(* IEC 61131-3 sources: esbmc-plc-benchmark-suite/ml/demo, 15 files *)

(* ---- airlock_door_interlock.st ---- *)
(* ============================================================
   Cleanroom airlock door interlock : demo program, not in the
   suite.
   Safety intent: the inner and outer airlock doors must never
   both be unlocked at the same time (maintains pressure
   differential and contamination control).
   ============================================================ *)
PROGRAM airlock_control
  VAR
    inner_request AT %IX0.0 : BOOL;
    outer_request AT %IX0.1 : BOOL;
    cycle_busy    AT %IX0.2 : BOOL;
    inner_unlocked AT %QX0.0 : BOOL;
    outer_unlocked AT %QX0.1 : BOOL;
  END_VAR

  IF NOT cycle_busy AND inner_request AND NOT outer_request THEN
    inner_unlocked := TRUE;
    outer_unlocked := FALSE;
  ELSIF NOT cycle_busy AND outer_request AND NOT inner_request THEN
    inner_unlocked := FALSE;
    outer_unlocked := TRUE;
  ELSE
    inner_unlocked := FALSE;
    outer_unlocked := FALSE;
  END_IF;
END_PROGRAM

CONFIGURATION Config0
  RESOURCE Res0 ON PLC
    TASK tcyclic(INTERVAL := T#10ms, PRIORITY := 0);
    PROGRAM inst0 WITH tcyclic : airlock_control;
  END_RESOURCE
END_CONFIGURATION

(* ---- burner_ignition.st ---- *)
(* ============================================================
   Gas burner ignition sequence : demo program, not in the suite.
   Safety intent: the gas valve must never open unless the purge
   fan has been confirmed running, and the spark igniter must
   never be energised while the gas valve is closed (no fuel to
   ignite, wasted spark risk is secondary to the interlock logic
   itself being sound).
   ============================================================ *)
PROGRAM burner_seq
  VAR
    purge_fan_ok  AT %IX0.0 : BOOL;
    start_request AT %IX0.1 : BOOL;
    flame_proven  AT %IX0.2 : BOOL;
    gas_valve     AT %QX0.0 : BOOL;
    igniter       AT %QX0.1 : BOOL;
  END_VAR

  IF start_request AND purge_fan_ok THEN
    gas_valve := TRUE;
  ELSE
    gas_valve := FALSE;
  END_IF;

  IF gas_valve AND NOT flame_proven THEN
    igniter := TRUE;
  ELSE
    igniter := FALSE;
  END_IF;
END_PROGRAM

CONFIGURATION Config0
  RESOURCE Res0 ON PLC
    TASK tcyclic(INTERVAL := T#10ms, PRIORITY := 0);
    PROGRAM inst0 WITH tcyclic : burner_seq;
  END_RESOURCE
END_CONFIGURATION

(* ---- conveyor_gate.st ---- *)
(* ============================================================
   Conveyor infeed gate : demo program, not in the benchmark suite.
   Safety intent: the infeed gate must never open while the
   downstream jam sensor is active, and the conveyor motor must
   never run while the gate is open (product would fall through).
   ============================================================ *)
PROGRAM gate_control
  VAR
    jam_sensor   AT %IX0.0 : BOOL;  (* downstream jam detected *)
    start_button AT %IX0.1 : BOOL;
    stop_button  AT %IX0.2 : BOOL;
    gate_open    AT %QX0.0 : BOOL;
    motor_run    AT %QX0.1 : BOOL;
  END_VAR

  IF stop_button OR jam_sensor THEN
    gate_open := FALSE;
    motor_run := FALSE;
  ELSIF start_button AND NOT jam_sensor THEN
    motor_run := TRUE;
  END_IF;

  IF motor_run THEN
    gate_open := FALSE;
  ELSE
    gate_open := TRUE;
  END_IF;
END_PROGRAM

CONFIGURATION Config0
  RESOURCE Res0 ON PLC
    TASK tcyclic(INTERVAL := T#10ms, PRIORITY := 0);
    PROGRAM inst0 WITH tcyclic : gate_control;
  END_RESOURCE
END_CONFIGURATION

(* ---- conveyor_with_distractor.st ---- *)
(* ============================================================
   Conveyor with unrelated diagnostic counter : demo program, not
   in the suite.
   Safety intent: the belt motor must never run while the
   emergency-stop rope switch is tripped. cycle_count is a
   diagnostic counter unrelated to any safety property.
   ============================================================ *)
PROGRAM belt_control
  VAR
    estop_tripped AT %IX0.0 : BOOL;
    run_request   AT %IX0.1 : BOOL;
    belt_motor    AT %QX0.0 : BOOL;
    cycle_count   : INT := 0;
  END_VAR

  IF estop_tripped THEN
    belt_motor := FALSE;
  ELSIF run_request THEN
    belt_motor := TRUE;
  END_IF;

  IF belt_motor THEN
    cycle_count := cycle_count + 1;
  END_IF;
END_PROGRAM

CONFIGURATION Config0
  RESOURCE Res0 ON PLC
    TASK tcyclic(INTERVAL := T#10ms, PRIORITY := 0);
    PROGRAM inst0 WITH tcyclic : belt_control;
  END_RESOURCE
END_CONFIGURATION

(* ---- door_interlock.st ---- *)
(* ============================================================
   Machine guard door interlock : demo program, not in the suite.
   Safety intent: the spindle must never run while the guard door
   is open.
   ============================================================ *)
PROGRAM guard_interlock
  VAR
    door_open    AT %IX0.0 : BOOL;
    start_button AT %IX0.1 : BOOL;
    spindle_run  AT %QX0.0 : BOOL;
  END_VAR

  IF door_open THEN
    spindle_run := FALSE;
  ELSIF start_button THEN
    spindle_run := TRUE;
  END_IF;
END_PROGRAM

CONFIGURATION Config0
  RESOURCE Res0 ON PLC
    TASK tcyclic(INTERVAL := T#10ms, PRIORITY := 0);
    PROGRAM inst0 WITH tcyclic : guard_interlock;
  END_RESOURCE
END_CONFIGURATION

(* ---- dual_heater.st ---- *)
(* ============================================================
   Dual immersion heater : demo program, not in the suite.
   Safety intent: heater_A and heater_B must never be energised
   together (shared circuit breaker is rated for one at a time).
   ============================================================ *)
PROGRAM dual_heater
  VAR
    demand_a  AT %IX0.0 : BOOL;
    demand_b  AT %IX0.1 : BOOL;
    heater_A  AT %QX0.0 : BOOL;
    heater_B  AT %QX0.1 : BOOL;
  END_VAR

  IF demand_a THEN
    heater_A := TRUE;
    heater_B := FALSE;
  ELSIF demand_b THEN
    heater_A := FALSE;
    heater_B := TRUE;
  ELSE
    heater_A := FALSE;
    heater_B := FALSE;
  END_IF;
END_PROGRAM

CONFIGURATION Config0
  RESOURCE Res0 ON PLC
    TASK tcyclic(INTERVAL := T#10ms, PRIORITY := 0);
    PROGRAM inst0 WITH tcyclic : dual_heater;
  END_RESOURCE
END_CONFIGURATION

(* ---- hoist_overload_cutoff.st ---- *)
(* ============================================================
   Crane hoist overload cutoff : demo program, not in the suite.
   Safety intent: the hoist motor must never raise the load while
   the overload sensor is tripped, regardless of the operator's
   raise command.
   ============================================================ *)
PROGRAM hoist_control
  VAR
    overload_tripped AT %IX0.0 : BOOL;
    raise_command    AT %IX0.1 : BOOL;
    lower_command    AT %IX0.2 : BOOL;
    hoist_raise       AT %QX0.0 : BOOL;
    hoist_lower       AT %QX0.1 : BOOL;
  END_VAR

  IF overload_tripped THEN
    hoist_raise := FALSE;
  ELSIF raise_command AND NOT lower_command THEN
    hoist_raise := TRUE;
  ELSE
    hoist_raise := FALSE;
  END_IF;

  hoist_lower := lower_command AND NOT raise_command;
END_PROGRAM

CONFIGURATION Config0
  RESOURCE Res0 ON PLC
    TASK tcyclic(INTERVAL := T#10ms, PRIORITY := 0);
    PROGRAM inst0 WITH tcyclic : hoist_control;
  END_RESOURCE
END_CONFIGURATION

(* ---- kiln_door_latch.st ---- *)
(* ============================================================
   Industrial kiln door safety latch : demo program, not in the
   suite.
   Safety intent: the heating element must never be energised
   while the kiln door is open; once the door has been opened
   during a heat cycle, the element stays locked out even after
   the door closes again, until an operator explicitly resets it.
   ============================================================ *)
PROGRAM kiln_control
  VAR
    door_open     AT %IX0.0 : BOOL;
    heat_request  AT %IX0.1 : BOOL;
    reset_button  AT %IX0.2 : BOOL;
    heater_element AT %QX0.0 : BOOL;
    door_fault_latched : BOOL := FALSE;
  END_VAR

  IF door_open THEN
    door_fault_latched := TRUE;
  ELSIF reset_button THEN
    door_fault_latched := FALSE;
  END_IF;

  IF door_fault_latched OR door_open THEN
    heater_element := FALSE;
  ELSIF heat_request THEN
    heater_element := TRUE;
  ELSE
    heater_element := FALSE;
  END_IF;
END_PROGRAM

CONFIGURATION Config0
  RESOURCE Res0 ON PLC
    TASK tcyclic(INTERVAL := T#10ms, PRIORITY := 0);
    PROGRAM inst0 WITH tcyclic : kiln_control;
  END_RESOURCE
END_CONFIGURATION

(* ---- press_two_hand.st ---- *)
(* ============================================================
   Hydraulic press two-hand safety control : demo program, not in
   the suite.
   Safety intent: the press ram must never descend unless both
   palm buttons are pressed simultaneously (prevents one-handed
   operation while the other hand is in the die area).
   ============================================================ *)
PROGRAM press_control
  VAR
    palm_left  AT %IX0.0 : BOOL;
    palm_right AT %IX0.1 : BOOL;
    light_curtain_clear AT %IX0.2 : BOOL;
    ram_descend AT %QX0.0 : BOOL;
  END_VAR

  IF palm_left AND palm_right AND light_curtain_clear THEN
    ram_descend := TRUE;
  ELSE
    ram_descend := FALSE;
  END_IF;
END_PROGRAM

CONFIGURATION Config0
  RESOURCE Res0 ON PLC
    TASK tcyclic(INTERVAL := T#10ms, PRIORITY := 0);
    PROGRAM inst0 WITH tcyclic : press_control;
  END_RESOURCE
END_CONFIGURATION

(* ---- pump_pressure_relief.st ---- *)
(* ============================================================
   Pump / pressure-relief valve : demo program, not in the
   benchmark suite.
   Safety intent: the feed pump must never run while the relief
   valve is closed (dead-heading risk), and the relief valve must
   never be closed while the high-pressure alarm is active.
   ============================================================ *)
PROGRAM pump_relief
  VAR
    hi_pressure_alarm AT %IX0.0 : BOOL;  (* pressure above safe limit *)
    pump_request      AT %IX0.1 : BOOL;
    manual_close       AT %IX0.2 : BOOL;
    pump_run          AT %QX0.0 : BOOL;
    relief_valve_open AT %QX0.1 : BOOL;
  END_VAR

  IF hi_pressure_alarm THEN
    relief_valve_open := TRUE;
  ELSIF manual_close AND NOT hi_pressure_alarm THEN
    relief_valve_open := FALSE;
  END_IF;

  IF relief_valve_open AND pump_request THEN
    pump_run := TRUE;
  ELSE
    pump_run := FALSE;
  END_IF;
END_PROGRAM

CONFIGURATION Config0
  RESOURCE Res0 ON PLC
    TASK tcyclic(INTERVAL := T#10ms, PRIORITY := 0);
    PROGRAM inst0 WITH tcyclic : pump_relief;
  END_RESOURCE
END_CONFIGURATION

(* ---- reactor_2oo3_trip.st ---- *)
(* ============================================================
   Reactor overpressure trip, 2-out-of-3 voting : demo program,
   not in the suite.
   Safety intent: the trip valve must open whenever at least two
   of the three independent pressure switches agree the vessel is
   over-pressured (2oo3 voting rejects a single sensor fault).
   ============================================================ *)
PROGRAM trip_2oo3
  VAR
    ps1 AT %IX0.0 : BOOL;
    ps2 AT %IX0.1 : BOOL;
    ps3 AT %IX0.2 : BOOL;
    trip_valve AT %QX0.0 : BOOL;
  END_VAR

  IF (ps1 AND ps2) OR (ps1 AND ps3) OR (ps2 AND ps3) THEN
    trip_valve := TRUE;
  ELSE
    trip_valve := FALSE;
  END_IF;
END_PROGRAM

CONFIGURATION Config0
  RESOURCE Res0 ON PLC
    TASK tcyclic(INTERVAL := T#10ms, PRIORITY := 0);
    PROGRAM inst0 WITH tcyclic : trip_2oo3;
  END_RESOURCE
END_CONFIGURATION

(* ---- silo_level.st ---- *)
(* ============================================================
   Grain silo fill control : demo program, not in the suite.
   Safety intent: the inlet auger must never run while the
   high-level sensor is tripped (overfill/structural risk), and
   the outlet gate must never open while the inlet auger runs
   (product would short-circuit straight through).
   ============================================================ *)
PROGRAM silo_fill
  VAR
    high_level    AT %IX0.0 : BOOL;
    fill_request  AT %IX0.1 : BOOL;
    empty_request AT %IX0.2 : BOOL;
    inlet_auger   AT %QX0.0 : BOOL;
    outlet_gate   AT %QX0.1 : BOOL;
  END_VAR

  IF high_level THEN
    inlet_auger := FALSE;
  ELSIF fill_request AND NOT empty_request THEN
    inlet_auger := TRUE;
  END_IF;

  IF inlet_auger THEN
    outlet_gate := FALSE;
  ELSIF empty_request THEN
    outlet_gate := TRUE;
  END_IF;
END_PROGRAM

CONFIGURATION Config0
  RESOURCE Res0 ON PLC
    TASK tcyclic(INTERVAL := T#10ms, PRIORITY := 0);
    PROGRAM inst0 WITH tcyclic : silo_fill;
  END_RESOURCE
END_CONFIGURATION

(* ---- three_pump_lockout.st ---- *)
(* ============================================================
   Three-pump station lockout : demo program, not in the suite.
   Safety intent: at most one of the three pumps may run at a time
   (shared discharge header cannot take combined flow).
   ============================================================ *)
PROGRAM three_pump
  VAR
    req_a AT %IX0.0 : BOOL;
    req_b AT %IX0.1 : BOOL;
    req_c AT %IX0.2 : BOOL;
    pump_a AT %QX0.0 : BOOL;
    pump_b AT %QX0.1 : BOOL;
    pump_c AT %QX0.2 : BOOL;
  END_VAR

  IF req_a THEN
    pump_a := TRUE;
    pump_b := FALSE;
    pump_c := FALSE;
  ELSIF req_b THEN
    pump_a := FALSE;
    pump_b := TRUE;
    pump_c := FALSE;
  ELSIF req_c THEN
    pump_a := FALSE;
    pump_b := FALSE;
    pump_c := TRUE;
  ELSE
    pump_a := FALSE;
    pump_b := FALSE;
    pump_c := FALSE;
  END_IF;
END_PROGRAM

CONFIGURATION Config0
  RESOURCE Res0 ON PLC
    TASK tcyclic(INTERVAL := T#10ms, PRIORITY := 0);
    PROGRAM inst0 WITH tcyclic : three_pump;
  END_RESOURCE
END_CONFIGURATION

(* ---- vent_fan_interlock.st ---- *)
(* ============================================================
   Paint booth vent fan / spray gun interlock : demo program, not
   in the suite.
   Safety intent: the spray gun trigger must be blocked whenever
   the exhaust fan is NOT running (solvent vapour must always be
   extracted while spraying).
   ============================================================ *)
PROGRAM booth_interlock
  VAR
    fan_running   AT %IX0.0 : BOOL;
    trigger_pull  AT %IX0.1 : BOOL;
    gun_enabled   AT %QX0.0 : BOOL;
  END_VAR

  IF NOT fan_running THEN
    gun_enabled := FALSE;
  ELSE
    gun_enabled := trigger_pull;
  END_IF;
END_PROGRAM

CONFIGURATION Config0
  RESOURCE Res0 ON PLC
    TASK tcyclic(INTERVAL := T#10ms, PRIORITY := 0);
    PROGRAM inst0 WITH tcyclic : booth_interlock;
  END_RESOURCE
END_CONFIGURATION

(* ---- welder_gas_shield.st ---- *)
(* ============================================================
   MIG welder shielding-gas interlock : demo program, not in the
   suite.
   Safety intent: the arc (weld current) must never strike unless
   BOTH the shielding-gas flow is confirmed AND the torch trigger
   is pulled; the arc must also be blocked whenever the gas flow
   sensor drops out mid-weld.
   ============================================================ *)
PROGRAM welder_control
  VAR
    gas_flow_ok   AT %IX0.0 : BOOL;
    trigger_pull  AT %IX0.1 : BOOL;
    arc_on        AT %QX0.0 : BOOL;
  END_VAR

  IF NOT gas_flow_ok THEN
    arc_on := FALSE;
  ELSIF trigger_pull AND gas_flow_ok THEN
    arc_on := TRUE;
  ELSE
    arc_on := FALSE;
  END_IF;
END_PROGRAM

CONFIGURATION Config0
  RESOURCE Res0 ON PLC
    TASK tcyclic(INTERVAL := T#10ms, PRIORITY := 0);
    PROGRAM inst0 WITH tcyclic : welder_control;
  END_RESOURCE
END_CONFIGURATION
